(* IEC 61131-3 sources: HypervisionPLC-SCADA/demo/vandvaerk, 3 files *)

(* ---- globals.st ---- *)
GLOBAL_VAR
  g_speed     : REAL;   (* L3: tidsfaktor 1-120 *)
  g_f_p1      : BOOL;   (* L3: broendpumpe fejl (scenarie 1) *)
  g_f_p2      : BOOL;   (* L3: doseringspumpe fejl *)
  g_f_an      : BOOL;   (* L3: analysatorfejl *)
  g_at2       : REAL;   (* L3: klor efter kontakttank mg/L, minus 1 = analysatorfejl *)
  g_well      : REAL;   (* L3: broendniveau m *)
  g_q         : REAL;   (* L3: flow l/s *)
  g_p1_run    : BOOL;   (* L3: broendpumpe koerer *)
  g_p2_run    : BOOL;   (* L3: doseringspumpe koerer *)
  g_xv1_open  : BOOL;   (* L3: skylleventil aaben *)
  g_hypo      : REAL;   (* L3: hypotank pct *)
  g_res       : REAL;   (* L3: hoejdebeholder pct *)
  g_vol       : REAL;   (* L3: doegnmaengde m3 *)
  g_p1_cmd    : BOOL;   (* L2: broendpumpe start *)
  g_p2_cmd    : BOOL;   (* L2: doseringspumpe start *)
  g_xv1_cmd   : BOOL;   (* L2: skylleventil aaben *)
  g_p2_pct    : REAL;   (* L2: doseringspumpens ydelse 0-100 pct *)
END_VAR

(* ---- logic2_styring.st ---- *)
PROGRAM VandvaerkStyring
(* Broendstation med klordosering, Logic2: styring. Driftsform (0 fra, 1 auto, 2 manuel), startsekvens (skyl,
   broendpumpe, dosering), stop, tilladelser, interlocks og alarmer. Dosering er flow-proportional med trim fra
   analysatoren efter kontakttanken. Ingen fysisk I/O. Interval 500 ms. Tider i sekunder paa den simulerede tid.
   VW_STATUS: 0 stoppet, 1 starter, 2 drift, 3 stopper, 4 trip.
   VW_TRIP: 0 ingen, 1 broend lav, 2 hypo eller dosering, 3 klor uden for graenser, 4 pumpe eller intet flow. *)
VAR
  VW_MODE        : INT := 1;
  VW_KVIT        : BOOL;
  VW_MAN_P1      : BOOL;
  VW_MAN_P2      : BOOL;
  VW_MAN_XV1     : BOOL;
  VW_SP_START    : REAL := 40.0;
  VW_SP_STOP     : REAL := 85.0;
  VW_SP_DOSE     : REAL := 1.0;
  VW_SP_RES      : REAL := 0.5;
  VW_TRIM        : BOOL := TRUE;
  VW_SP_LAV      : REAL := 0.2;
  VW_SP_HOEJ     : REAL := 2.0;
  VW_STATUS      : INT;
  VW_TRIN        : INT;
  VW_TRIP        : INT;
  VW_KOM_P1      : BOOL;
  VW_KOM_P2      : BOOL;
  VW_KOM_XV1     : BOOL;
  VW_DOSIS_EFF   : REAL := 1.0;
  VW_P2_PCT      : REAL;
  VW_ALARMER     : INT;
  VW_AL_BROND    : BOOL;
  VW_AL_BROND_LL : BOOL;
  VW_AL_HYPO     : BOOL;
  VW_AL_HYPO_TOM : BOOL;
  VW_AL_KLOR_LAV : BOOL;
  VW_AL_KLOR_HOEJ: BOOL;
  VW_AL_P1       : BOOL;
  VW_AL_P2       : BOOL;
  VW_AL_FLOW     : BOOL;
  VW_AL_DOEGN    : BOOL;
  VW_AL_AN       : BOOL;
  VW_AL_BEH_LAV  : BOOL;
  VW_AL_BEH_HOEJ : BOOL;
  VW_AL_TRIP     : BOOL;
  trin           : INT;
  trip           : BOOL;
  trip_now       : INT;
  want           : BOOL;
  perm           : BOOL;
  permrun        : BOOL;
  clvalid        : BOOL;
  ack            : BOOL;
  p1             : BOOL;
  p2             : BOOL;
  xv1            : BOOL;
  t_step         : REAL;
  t_run          : REAL;
  t_hi           : REAL;
  t_lo           : REAL;
  t_nf           : REAL;
  t_nd           : REAL;
  dt             : REAL;
END_VAR
BEGIN
  dt := 0.5 * MAX(g_speed, 1.0);
  VW_MODE := LIMIT(0, VW_MODE, 2);
  ack := VW_KVIT;
  VW_KVIT := FALSE;
  clvalid := (NOT g_f_an) AND (g_at2 >= 0.0);

  (* tilladelser: til at starte, og til at blive ved at koere *)
  perm := (g_well >= 3.0) AND (g_hypo >= 10.0) AND (NOT g_f_p1) AND (NOT g_f_p2) AND (g_vol < 2400.0) AND (NOT trip);
  permrun := (g_well >= 1.5) AND (g_hypo >= 5.0) AND (g_res < 97.0) AND (g_vol < 2400.0);

  (* timere til interlocks: klor i simuleret tid, hardware i rigtig tid (0,5 s pr. scan) *)
  IF g_p2_run THEN t_run := t_run + dt; ELSE t_run := 0.0; END_IF;
  IF clvalid AND (g_q > 1.0) AND (g_at2 > VW_SP_HOEJ) THEN t_hi := t_hi + dt; ELSE t_hi := 0.0; END_IF;
  IF clvalid AND g_p2_run AND (t_run >= 900.0) AND (g_at2 < VW_SP_LAV) THEN t_lo := t_lo + dt; ELSE t_lo := 0.0; END_IF;
  IF g_p1_cmd AND (g_q < 10.0) THEN t_nf := t_nf + 0.5; ELSE t_nf := 0.0; END_IF;
  IF g_p2_cmd AND (NOT g_p2_run) THEN t_nd := t_nd + 0.5; ELSE t_nd := 0.0; END_IF;

  (* trip: groeft aarsag i prioriteret raekkefoelge, laast til kvittering naar aarsagen er vaek *)
  trip_now := 0;
  IF g_p1_cmd AND (g_well < 1.0) THEN
    trip_now := 1;
  ELSIF g_p2_cmd AND ((g_hypo < 3.0) OR (t_nd >= 10.0)) THEN
    trip_now := 2;
  ELSIF (t_hi >= 30.0) OR (t_lo >= 600.0) THEN
    trip_now := 3;
  ELSIF (g_p1_cmd AND g_f_p1) OR (t_nf >= 20.0) THEN
    trip_now := 4;
  END_IF;
  IF (trip_now > 0) AND (NOT trip) THEN
    trip := TRUE;
    VW_TRIP := trip_now;
  END_IF;
  IF trip AND ack AND (trip_now = 0) THEN
    trip := FALSE;
    VW_TRIP := 0;
  END_IF;

  (* oensket drift i auto: niveau i hoejdebeholderen med hysterese *)
  IF VW_MODE = 1 THEN
    IF g_res <= VW_SP_START THEN want := TRUE; END_IF;
    IF g_res >= VW_SP_STOP THEN want := FALSE; END_IF;
  ELSE
    want := FALSE;
  END_IF;

  IF trip THEN
    trin := 0;
    p1 := FALSE;
    p2 := FALSE;
    xv1 := FALSE;
  ELSIF VW_MODE = 2 THEN
    (* manuel: interlocks gaelder stadig *)
    trin := 0;
    p1 := VW_MAN_P1 AND (g_well >= 1.5) AND (NOT g_f_p1);
    p2 := VW_MAN_P2 AND g_p1_run AND (g_hypo >= 3.0);
    xv1 := VW_MAN_XV1 AND (NOT p1);
  ELSIF trin = 0 THEN
    p1 := FALSE;
    p2 := FALSE;
    xv1 := FALSE;
    IF want AND perm THEN
      trin := 1;
      t_step := 0.0;
    END_IF;
  ELSIF trin = 1 THEN
    (* skyl: skylleventilen aaben i 30 s *)
    xv1 := TRUE;
    t_step := t_step + dt;
    IF (NOT want) OR (NOT permrun) THEN
      trin := 5;
      t_step := 0.0;
    ELSIF g_xv1_open AND (t_step >= 30.0) THEN
      trin := 2;
      t_step := 0.0;
    END_IF;
  ELSIF trin = 2 THEN
    (* broendpumpen starter, skylleventilen lukker, vent paa stabilt flow *)
    xv1 := FALSE;
    p1 := TRUE;
    t_step := t_step + dt;
    IF (NOT want) OR (NOT permrun) THEN
      trin := 5;
      t_step := 0.0;
    ELSIF (g_q >= 20.0) AND (t_step >= 15.0) THEN
      trin := 3;
      t_step := 0.0;
    END_IF;
  ELSIF trin = 3 THEN
    (* dosering starter *)
    p2 := TRUE;
    t_step := t_step + dt;
    IF (NOT want) OR (NOT permrun) THEN
      trin := 5;
      t_step := 0.0;
    ELSIF g_p2_run AND (t_step >= 10.0) THEN
      trin := 4;
      t_step := 0.0;
    END_IF;
  ELSIF trin = 4 THEN
    IF (NOT want) OR (NOT permrun) THEN
      trin := 5;
      t_step := 0.0;
    END_IF;
  ELSE
    (* stop: doseringen foerst, saa broendpumpen *)
    p2 := FALSE;
    t_step := t_step + dt;
    IF t_step >= 10.0 THEN p1 := FALSE; END_IF;
    IF t_step >= 20.0 THEN trin := 0; END_IF;
  END_IF;

  (* flow-proportional dosering: l/t = flow l/s * dosis mg/l * 3600 / 120000 (12 pct hypo er 120 g/l); trim fra AT2 *)
  IF VW_TRIM AND clvalid AND (t_run >= 900.0) THEN
    VW_DOSIS_EFF := LIMIT(0.2, VW_SP_DOSE + 0.5 * (VW_SP_RES - g_at2), 3.0);
  ELSE
    VW_DOSIS_EFF := VW_SP_DOSE;
  END_IF;
  VW_P2_PCT := LIMIT(0.0, g_q * VW_DOSIS_EFF * 0.03 / 5.0 * 100.0, 100.0);
  g_p2_pct := VW_P2_PCT;

  g_p1_cmd := p1;
  g_p2_cmd := p2;
  g_xv1_cmd := xv1;
  VW_KOM_P1 := p1;
  VW_KOM_P2 := p2;
  VW_KOM_XV1 := xv1;
  VW_TRIN := trin;

  IF trip THEN
    VW_STATUS := 4;
  ELSIF trin = 5 THEN
    VW_STATUS := 3;
  ELSIF (trin >= 1) AND (trin <= 3) THEN
    VW_STATUS := 1;
  ELSIF (trin = 4) OR (g_p1_run AND (VW_MODE = 2)) THEN
    VW_STATUS := 2;
  ELSE
    VW_STATUS := 0;
  END_IF;

  VW_AL_BROND := g_well < 2.0;
  VW_AL_BROND_LL := g_well < 1.0;
  VW_AL_HYPO := g_hypo < 15.0;
  VW_AL_HYPO_TOM := g_hypo < 3.0;
  VW_AL_KLOR_LAV := t_lo >= 120.0;
  VW_AL_KLOR_HOEJ := clvalid AND (g_at2 > VW_SP_HOEJ);
  VW_AL_P1 := g_f_p1;
  VW_AL_P2 := g_f_p2;
  VW_AL_FLOW := t_nf >= 10.0;
  VW_AL_DOEGN := g_vol > 2160.0;
  VW_AL_AN := g_f_an;
  VW_AL_BEH_LAV := g_res < 20.0;
  VW_AL_BEH_HOEJ := g_res > 95.0;
  VW_AL_TRIP := trip;
  VW_ALARMER := BOOL_TO_INT(VW_AL_BROND) + BOOL_TO_INT(VW_AL_BROND_LL) + BOOL_TO_INT(VW_AL_HYPO) + BOOL_TO_INT(VW_AL_HYPO_TOM)
              + BOOL_TO_INT(VW_AL_KLOR_LAV) + BOOL_TO_INT(VW_AL_KLOR_HOEJ) + BOOL_TO_INT(VW_AL_P1) + BOOL_TO_INT(VW_AL_P2)
              + BOOL_TO_INT(VW_AL_FLOW) + BOOL_TO_INT(VW_AL_DOEGN) + BOOL_TO_INT(VW_AL_AN) + BOOL_TO_INT(VW_AL_BEH_LAV)
              + BOOL_TO_INT(VW_AL_BEH_HOEJ) + BOOL_TO_INT(VW_AL_TRIP);
END_PROGRAM

(* ---- logic3_proces.st ---- *)
PROGRAM VandvaerkProces
(* Broendstation med klordosering, Logic3: procesmodel. Broend med tilstroemning fra grundvandet, broendpumpe
   (35 l/s, 10 s opstart), trykmaaler, skylleventil (8 s gangtid), hypotank (50 l) med doseringspumpe (5 l/t),
   hoejdebeholder (300 m3) med doegnets forbrug og doegnmaengde. Klor: doseret koncentration (mg/l) = doseret
   hypo l/t * 120000 / flow l/t (12 pct hypo er 120 g/l). AT1 er efter indsproejtningen, AT2 efter kontakttanken
   (40 m3, 1. ordens forsinkelse med V / flow og lille nedbrydning). CT er klor gange kontakttid. Klokke,
   tidsfaktor og scenarier. Interval 500 ms.
   VW_SCEN: 0 normal, 1 broendpumpe fejl, 2 hypotank tom, 3 hoej efterspoergsel (2,5 gange), 4 overdosering (4 gange).
   Fejl der kan kombineres: VW_F_AN analysatorfejl, VW_F_P2 doseringspumpe fejl, VW_F_LAV lav grundvandsstand. *)
VAR
  VW_SPEED      : REAL := 10.0;
  VW_SCEN       : INT;
  VW_F_AN       : BOOL;
  VW_F_P2       : BOOL;
  VW_F_LAV      : BOOL;
  VW_KLOKKE     : REAL;
  VW_BROND      : REAL := 8.0;
  VW_Q          : REAL;
  VW_TRYK       : REAL;
  VW_P1_FB      : BOOL;
  VW_XV1_AABEN  : BOOL;
  VW_XV1_LUKKET : BOOL := TRUE;
  VW_XV1_POS    : REAL;
  VW_P2_FB      : BOOL;
  VW_FYLD       : BOOL;
  VW_HYPO       : REAL := 90.0;
  VW_P2_LH      : REAL;
  VW_BEH        : REAL := 35.0;
  VW_BEHOV      : REAL;
  VW_DOEGN      : REAL;
  VW_DOSE       : REAL;
  VW_AT1        : REAL;
  VW_AT2        : REAL;
  VW_TKONT      : REAL;
  VW_CT         : REAL;
  t_dag         : REAL := 21600.0;
  f_p1          : BOOL;
  over          : BOOL;
  dem_x         : REAL := 1.0;
  rech_x        : REAL := 1.0;
  ramp          : REAL;
  rech          : REAL;
  luft          : REAL;
  c1            : REAL;
  c2            : REAL;
  tau           : REAL;
  dt            : REAL;
  last_hour     : REAL;
END_VAR
BEGIN
  VW_SPEED := LIMIT(1.0, VW_SPEED, 120.0);
  g_speed := VW_SPEED;
  dt := 0.5 * VW_SPEED;

  (* klokken starter kl. 6 og gaar rundt i doegn *)
  t_dag := t_dag + dt;
  IF t_dag >= 86400.0 THEN t_dag := t_dag - 86400.0; END_IF;
  VW_KLOKKE := t_dag / 3600.0;

  (* scenarier og fejl *)
  VW_SCEN := LIMIT(0, VW_SCEN, 4);
  f_p1 := (VW_SCEN = 1);
  over := (VW_SCEN = 4);
  IF VW_SCEN = 3 THEN dem_x := 2.5; ELSE dem_x := 1.0; END_IF;
  IF VW_F_LAV THEN rech_x := 0.3; ELSE rech_x := 1.0; END_IF;
  g_f_p1 := f_p1;
  g_f_p2 := VW_F_P2;
  g_f_an := VW_F_AN;

  (* broendpumpen: 10 s op, 6 s ned; trukket tom for vand falder ydelsen *)
  IF g_p1_cmd AND (NOT f_p1) THEN
    ramp := MIN(1.0, ramp + dt / 10.0);
  ELSE
    ramp := MAX(0.0, ramp - dt / 6.0);
  END_IF;
  VW_P1_FB := ramp > 0.5;
  luft := LIMIT(0.0, (VW_BROND - 0.3) / 0.7, 1.0);
  VW_Q := 35.0 * ramp * luft;
  rech := 70.0 * rech_x * (10.0 - VW_BROND) / 10.0;
  VW_BROND := LIMIT(0.0, VW_BROND + (rech - VW_Q) * dt / 3000.0, 10.0);
  VW_TRYK := ramp * (3.0 + 0.02 * VW_BEH);

  (* skylleventil: 8 s gangtid *)
  IF g_xv1_cmd THEN
    VW_XV1_POS := MIN(100.0, VW_XV1_POS + dt / 8.0 * 100.0);
  ELSE
    VW_XV1_POS := MAX(0.0, VW_XV1_POS - dt / 8.0 * 100.0);
  END_IF;
  VW_XV1_AABEN := VW_XV1_POS >= 95.0;
  VW_XV1_LUKKET := VW_XV1_POS <= 5.0;

  (* hypo: doseringspumpen kan give 5 l/t; overdosering er 4 gange; tanken er 50 l *)
  VW_P2_FB := g_p2_cmd AND (NOT VW_F_P2);
  IF VW_P2_FB THEN
    VW_P2_LH := 5.0 * g_p2_pct / 100.0;
    IF over THEN VW_P2_LH := VW_P2_LH * 4.0; END_IF;
  ELSE
    VW_P2_LH := 0.0;
  END_IF;
  IF VW_FYLD THEN
    VW_HYPO := 100.0;
    VW_FYLD := FALSE;
  END_IF;
  VW_HYPO := LIMIT(0.0, VW_HYPO - VW_P2_LH * dt / 3600.0 / 50.0 * 100.0, 100.0);
  IF VW_SCEN = 2 THEN VW_HYPO := MIN(VW_HYPO, 2.0); END_IF;

  (* forbrug: 20 l/s i middel, mest om eftermiddagen; hoejdebeholderen er 300 m3 *)
  VW_BEHOV := 20.0 * (1.0 + 0.6 * SIN(6.2832 * (VW_KLOKKE - 9.0) / 24.0)) * dem_x;
  VW_BEH := LIMIT(0.0, VW_BEH + (VW_Q - VW_BEHOV) * dt / 1000.0 / 300.0 * 100.0, 100.0);

  (* doegnmaengde nulstilles ved midnat *)
  VW_DOEGN := VW_DOEGN + VW_Q * dt / 1000.0;
  IF VW_KLOKKE < last_hour THEN VW_DOEGN := 0.0; END_IF;
  last_hour := VW_KLOKKE;

  (* klor: doseret koncentration, blanding, kontakttank *)
  IF VW_Q > 0.5 THEN
    VW_DOSE := VW_P2_LH * 120000.0 / (VW_Q * 3600.0);
  ELSE
    VW_DOSE := 0.0;
  END_IF;
  c1 := c1 + (VW_DOSE - c1) * MIN(1.0, dt / 20.0);
  IF VW_Q > 1.0 THEN
    tau := 40000.0 / VW_Q;
    VW_TKONT := MIN(40000.0 / VW_Q / 60.0, 999.0);
  ELSE
    tau := 1000000.0;
    VW_TKONT := 0.0;
  END_IF;
  c2 := MAX(0.0, c2 + ((c1 - c2) / tau - 0.00005 * c2) * dt);
  VW_AT1 := c1;
  IF VW_F_AN THEN
    VW_AT2 := -1.0;
    VW_CT := 0.0;
  ELSE
    VW_AT2 := c2;
    VW_CT := c2 * VW_TKONT;
  END_IF;

  g_at2 := VW_AT2;
  g_well := VW_BROND;
  g_q := VW_Q;
  g_p1_run := VW_P1_FB;
  g_p2_run := VW_P2_FB;
  g_xv1_open := VW_XV1_AABEN;
  g_hypo := VW_HYPO;
  g_res := VW_BEH;
  g_vol := VW_DOEGN;
END_PROGRAM
